(* IEC 61131-3 sources: SRCI_CLIENT_PLC/RobotLibrary/Library/POUs/Read/MC_ReadToolData/Structures, 4 files *)

(* ---- ReadToolDataOutCmd.st ---- *)
{attribute 'pack_mode' := '1'}
// -------------------------------------------------------------------------
//  SRCI Robot Library
// -------------------------------------------------------------------------
//
//  Object:      ReadToolDataOutCmd
//  Author:      Thorsten Brach
//  Date:        2024-08-09
//
//  Description:
//
//
//  Copyright:
//    (C) 2024 Thorsten Brach. All rights reserved
//             Licensed under the MIT License.
//
//  Disclaimer:
//    This project is provided without any guarantee and can be used for
//    private and commercial purposes. Any use is at the user’s
//    own risk and responsibility.
//
// -------------------------------------------------------------------------
TYPE ReadToolDataOutCmd :
STRUCT
  /// Tool index
  ToolNoReturn       : USINT;
  /// Tool data (see chapter 5.5.6.3)
  ToolData           : ToolData;
END_STRUCT
END_TYPE

(* ---- ReadToolDataParCmd.st ---- *)
{attribute 'pack_mode' := '1'}
// -------------------------------------------------------------------------
//  SRCI Robot Library
// -------------------------------------------------------------------------
//
//  Object:      ReadToolDataParCmd
//  Author:      Thorsten Brach
//  Date:        2024-08-09
//
//  Description:
//
//
//  Copyright:
//    (C) 2024 Thorsten Brach. All rights reserved
//             Licensed under the MIT License.
//
//  Disclaimer:
//    This project is provided without any guarantee and can be used for
//    private and commercial purposes. Any use is at the user’s
//    own risk and responsibility.
//
// -------------------------------------------------------------------------
TYPE ReadToolDataParCmd :
STRUCT
  /// Tool index
  /// • -1: Currently used tool on RC
  /// •  0: Flange -  Not possible to change
  /// • 1 (default)..254: Tool Frame
  ToolNo             : INT := 1; // ST-FIX F156: spec 6.2.17: '1 (default)'
END_STRUCT
END_TYPE

(* ---- ReadToolDataRecvData.st ---- *)
{attribute 'pack_mode' := '1'}
// -------------------------------------------------------------------------
//  SRCI Robot Library
// -------------------------------------------------------------------------
//
//  Object:      ReadToolDataRecvData
//  Author:      Thorsten Brach
//  Date:        2024-08-09
//
//  Description:
//
//
//  Copyright:
//    (C) 2024 Thorsten Brach. All rights reserved
//             Licensed under the MIT License.
//
//  Disclaimer:
//    This project is provided without any guarantee and can be used for
//    private and commercial purposes. Any use is at the user’s
//    own risk and responsibility.
//
// -------------------------------------------------------------------------
TYPE ReadToolDataRecvData EXTENDS RspHeader :
STRUCT
  /// Reserve
  Reserve       : BYTE;
  /// Tool index
  ToolNoReturn  : USINT;
  /// Tool data (see chapter 5.5.6.3)
  ToolData      : ToolData;
  /// The status bit "DataChanged" represents the modification state
  DataChanged   : BOOL;
END_STRUCT
END_TYPE

(* ---- ReadToolDataSendData.st ---- *)
{attribute 'pack_mode' := '1'}
// -------------------------------------------------------------------------
//  SRCI Robot Library
// -------------------------------------------------------------------------
//
//  Object:      ReadToolDataSendData
//  Author:      Thorsten Brach
//  Date:        2024-08-09
//
//  Description:
//
//
//  Copyright:
//    (C) 2024 Thorsten Brach. All rights reserved
//             Licensed under the MIT License.
//
//  Disclaimer:
//    This project is provided without any guarantee and can be used for
//    private and commercial purposes. Any use is at the user’s
//    own risk and responsibility.
//
// -------------------------------------------------------------------------
TYPE ReadToolDataSendData EXTENDS CmdHeader:
STRUCT
  /// Tool index
  /// • -1: Currently used tool on RC
  /// •  0: Flange -  Not possible to change
  /// • 1 (default)..254: Tool Frame
  ToolNo             : USINT;
END_STRUCT
END_TYPE
